Staubli VAL3: HMI_IO.dtx

mdesc mNomSpeed
num nPage
num nPageIndex
num nItemIndex
public bool bBool[11]
public string sUsingBus
bool bComment[16]
public string sLabel[16]
num nShowPageIndex
string sShowPageIndex
string sPageNum
public string sComment[16]
num nType
num nSelType
bool bRefresh
public string sValue[16]
bool bBtnHidden
bool bLabelHidden
num _nClock
bool bBack
num nDigCount
num nAngCount
bool bConfirm
bool bCancel
